(* IEC 61131-3 sources: Test002/ConveyorBelt/Class/VaranManager (part 2) *)

      7 : // all Varan_Base are ready with init
          if (s_ModuleList.ud_NrOfModules = 0) & (bEnableManagerWithNoModules = FALSE) then
            // penultimate call: if there are no clients => tell the hwcontrol to disable this
            To_HwControl.DisableVaranManager( ud_manager_number := VaranManagerNr
                                            , p_function_list   := #s_VMFunctions
                                            );
            State 		:= _NotInitialized;
          	ManagerOn := 0;                   //Disables Rt Task
          	bDisableCyTaskNoModules := TRUE;  //Disables Cy Task
          end_if;

    end_case;

    //trigger watchdog in init
    TriggerWatchdog();

  end_if;

  //increment our initcounter
  s_VaranManagerSettings.us_InitCounter += 1;

END_FUNCTION //VIRTUAL GLOBAL VaranManager::Init

//[#ENGLISH]
//=================================================================================================
//This function is called in PostScan by VaranManagerPostScan
//=================================================================================================
//[servers]	ManagerOn				:R		:state of Manager (On/Off)
//			RetryCounter			:W		:server counts retries
//			AsyVaranTime			:W		:time of asynchronous varan task
//[members]	s_CyHandles				:R		:structure to save Handles and thisp for cyclic update methodes
//			s_VaranTimes			:W		:structure for varan time measurement
//			us_UpdateOkCy			:R/W	:if variable = 1 then varan classes are called
//			p_ManagerStructure		:R		:pointer for manager structure (from OS)
//			s_VaranManagerSettings	:R/W	:structure for different varan settings
FUNCTION VIRTUAL GLOBAL VaranManager::CyWork
  VAR_INPUT
    EAX		              : UDINT;
  END_VAR
  VAR_OUTPUT
    state	    	        : UDINT;
  END_VAR
  VAR
    us_retry_counter	  : USINT;
    pHelp               : ^t_s_OneHandle;
    asyState            : UDINT;
    asyTimestamp        : UDINT;
  #ifndef VARAN_TIME_MEASUREMENT_DEACTIVATE
    ud_time				      : UDINT;
  #endif
    i				          	: UDINT;
    AsyReady            : BOOL;
    pHelpPostInit       : ^t_s_PostInitList;
  #ifdef VARAN_TIME_MEASUREMENT_SINGLE_OBJECTS
    ud_SingleTimeMark1  : UDINT;
    ud_SingleTimeMark2  : UDINT;
  #endif
  END_VAR

  //look if structur is ok, also check if cywork should be disabled due to no connected modules
  if ( p_ManagerStructure = NIL & b_PayloadSupport = false) | ( bDisableCyTaskNoModules = TRUE ) then
    return;
  end_if;

  //look if cyclic task is ready (executed)
  if b_PayloadSupport &
     pMultiVaran^.udVersion >= VM_MULTIVARAN_DOL_TIMING_AVAILABLE then

    MULTI_VARAN_iGetNodeProperty( hNodeHandle       := vmNodeHandle
                                , udPropertyId      := VM_PROP_TASK_STATE_ASY
                                , pudPropertyValue  := #asyState
                                );

    if asyState = TK_STATE_EXECUTING then
      AsyReady := FALSE;
    else
      AsyReady := TRUE;
    end_if;
  else
    AsyReady := (p_ManagerStructure^.sASY.ucHandshake and 16#10 ) <> 0;
  end_if;

#ifdef _LSL_TARGETARCH_ARM  // IO Image only needed for ARM  CPUs
#ifdef VARAN_iGetInputImage
  //look if manager is on or we are in post init phase (ManagerOn will be set in first realtime but we want to do something here in postinit)
  if ( ManagerOn = 1 ) | bPostInitActive = TRUE then
    if AsyReady then
      if b_IOImage then
        VARAN_iGetInputImage(VaranManagerNr, VARAN_DOL_ASY);
      end_if;
    end_if;
  end_if;
#endif
#endif

  // if there is a safety manager, we have to call it (but not from post init)
  if SafetyManagerThis & (bPostInitActive = FALSE) then
    SafetyManagerThis^.CyWork(0);
  end_if;

  //------------------------------------------------------------------------------------------------
  //first check Error
  if ( s_VaranManagerSettings.b_LogError = TRUE ) then
    LogError();
  end_if;

  // then check for rt log
  if bd_RtLog then
    if bd_RtLog.WatchdogTriggerFailed & (bd_RtLogged.WatchdogTriggerFailed = FALSE) then
#ifdef HWC_LogError
    HWC_LogError(this, "@0022 (VaranManager::CyWork) [SL] Error triggering the VaranManager Watchdog!");
#endif

      bd_RtLogged.WatchdogTriggerFailed := TRUE;
    end_if;

    if bd_RtLog.TimeSliceError & (bd_RtLogged.TimeSliceError = FALSE) then
#ifdef HWC_LogError
      HWC_LogError(this,"@019A (VaranManager::CyWork) Timeslice Error! Manager is set off!");
#endif

      bd_RtLogged.TimeSliceError := TRUE;
    end_if;

    bd_RtLog := 0;
  end_if;

#ifndef VARAN_TIME_MEASUREMENT_DEACTIVATE
  //measure time for cyclic
  ud_time := GetNsTime();
  s_VaranTimes.s_Cyclic.ud_CallTime := ( ud_time - s_VaranTimes.s_Cyclic.ud_Timemark ) / 1000;
  s_VaranTimes.s_Cyclic.ud_Timemark := ud_time;
#endif

  //check if we must disable a device
  if ( b_Disabledevice = TRUE ) then
    DisableDevice();
  end_if;

  //Update retry Counter
  if b_PayloadSupport &
     pMultiVaran^.udVersion >= VM_MULTIVARAN_VERSION_FULL_PAYLOAD_AVAILABLE  then
    MULTI_VARAN_iGetNodeProperty( hNodeHandle       := vmNodeHandle
                                , udPropertyId      := VM_PROP_GLOBAL_FAILED_ACCESS_COUNTER
                                , pudPropertyValue  := (#us_retry_counter)$^UDINT
                                );
  else
    us_retry_counter := p_ManagerStructure^.ucGlobalretryCounter;
  end_if;

  //look for change
  if ( us_retry_counter <> s_VaranManagerSettings.us_OldRetryCounter ) then

    //save on global counter
    RetryCounter += TO_USINT( us_retry_counter - s_VaranManagerSettings.us_OldRetryCounter );

    //save new counter
    s_VaranManagerSettings.us_OldRetryCounter := us_retry_counter;

    //update module retry counters cyclic
    if ( s_CyHandles.ud_NrOfHandles > 0 ) then

      //call all connected classes
      pHelp := #s_CyHandles.p_HandleList^[0];
      for i := 0 to s_CyHandles.ud_NrOfHandles - 1 do

        //call class
        pHelp^.p_This^.UpdateRetryCounter();

        //get pointer on next handle
        pHelp += sizeof(t_s_OneHandle);
      end_for;
    end_if;

    //update module retry counters cyclic
    if ( s_RtHandles.ud_NrOfHandles > 0 ) then

      //call all connected classes
      pHelp := #s_RtHandles.p_HandleList^[0];
      for i := 0 to s_RtHandles.ud_NrOfHandles - 1 do

        //call class
        pHelp^.p_This^.UpdateRetryCounter();

        //get pointer on next handle
        pHelp += sizeof(t_s_OneHandle);
      end_for;
    end_if;
  end_if;

  //look if manager is on or we are in post init phase (ManagerOn will be set in first realtime but we want to do something here in postinit)
  if ( ManagerOn = 1 ) | bPostInitActive = TRUE then

    //------------------------------------------------------------------------------------------------
    //look if cyclic task is ready (executed)
    if AsyReady = FALSE then
      s_VaranManagerSettings.us_NoCyclicUpdateCnt += 1;
      return;
    end_if;

#ifndef VARAN_TIME_MEASUREMENT_DEACTIVATE
    //------------------------------------------------------------------------------------------------
    //calculate cyclictime of varan task
    if b_PayloadSupport &
       pMultiVaran^.udVersion >= VM_MULTIVARAN_VERSION_FULL_PAYLOAD_AVAILABLE  then
      MULTI_VARAN_iGetNodeProperty( hNodeHandle       := vmNodeHandle
                                  , udPropertyId      := VM_PROP_ASY_TIME_UP_COUNTER
                                  , pudPropertyValue  := #asyTimestamp
                                  );
    else
      asyTimestamp := p_ManagerStructure^.sASY.uiTTUpCounter;
    end_if;

    if ( s_VaranTimes.s_AsyVaranTime.us_NotFirstRun	= 0 ) then

      //get counter of asy task
      s_VaranTimes.s_AsyVaranTime.ud_Timestamp := asyTimestamp;

      //start asy task
      if ( s_CyHandles.b_ExecuteDOL = TRUE ) then
        ExecuteDOL( VARAN_DOL_ASY );
      end_if;

      s_VaranTimes.s_AsyVaranTime.us_NotFirstRun := 1;
      return;
    end_if;

    //calculate ASY Time
    s_VaranTimes.s_AsyVaranTime.ud_ActUsageRate := asyTimestamp - s_VaranTimes.s_AsyVaranTime.ud_Timestamp;
    s_VaranTimes.s_AsyVaranTime.ud_Timestamp    := asyTimestamp;

    //look for maximum value
    if ( s_VaranTimes.s_AsyVaranTime.ud_ActUsageRate > s_VaranTimes.s_AsyVaranTime.ud_MaxUsageRate ) then
      s_VaranTimes.s_AsyVaranTime.ud_MaxUsageRate := s_VaranTimes.s_AsyVaranTime.ud_ActUsageRate;
    end_if;

    //save on server
    AsyVaranTime$UDINT := s_VaranTimes.s_AsyVaranTime.ud_ActUsageRate;
#endif

    //----------------------------------------------------------------------------------------------
    //hardware class handling

    // in post init we call only the modules which are logged in for post init
    if bPostInitActive then
      if PostInitModuleCnt then
        pHelpPostInit := #aPostInitList[0];
        for i := 0 to PostInitModuleCnt - 1 do

          //call class, if it's still not ready
          if pHelpPostInit^.p_This & pHelpPostInit^.b_CallMe then
            pHelpPostInit^.p_This^.UpdateCy();
          end_if;

          // set pointer on next this pointer
          pHelpPostInit += sizeof(t_s_PostInitList);
        end_for;
      end_if;
    else
      //look if we have classes
      if ( s_CyHandles.ud_NrOfHandles > 0 ) then

        //call all connected classes
        pHelp := #s_CyHandles.p_HandleList^[0];
        for i := 0 to s_CyHandles.ud_NrOfHandles - 1 do

#ifdef VARAN_TIME_MEASUREMENT_SINGLE_OBJECTS
          ud_SingleTimeMark1 := OS_READMICROSEC();
#endif

          //call class
          pHelp^.p_This^.UpdateCy();

#ifdef VARAN_TIME_MEASUREMENT_SINGLE_OBJECTS
          ud_SingleTimeMark2 := OS_READMICROSEC();
          pHelp^.TimeMeasuring.ud_ActTime := ud_SingleTimeMark2 - ud_SingleTimeMark1;

          if pHelp^.TimeMeasuring.ud_ActTime > pHelp^.TimeMeasuring.ud_MaxTime then
            pHelp^.TimeMeasuring.ud_MaxTime := pHelp^.TimeMeasuring.ud_ActTime;
          end_if;

          if pHelp^.TimeMeasuring.ud_ActTime < pHelp^.TimeMeasuring.ud_MinTime then
            pHelp^.TimeMeasuring.ud_MinTime := pHelp^.TimeMeasuring.ud_ActTime;
          end_if;
#endif

          //get pointer on next handle
          pHelp += sizeof(t_s_OneHandle);
        end_for;
      end_if;
    end_if;

    //start asy task
    if ( s_CyHandles.b_ExecuteDOL = TRUE ) then
      ExecuteDOL( VARAN_DOL_ASY );
    end_if;

  //------------------------------------------------------------ Client Instructions --------------------------------------------------------|
  //                                                                                                                                         V
    //DPRAM data handling
    if ( IsAlsoClient & p_ManagerClientSpace <> NIL ) then

      // copy data to ram
      // ->WRITE<-
      To_Stdlib.MemCpy( dest := #p_ASYDataWrite^.a_Data[0],     // Mem for p_ASYDataWrite is reserved in VaranManager2
                        source := AsyWriteData.pSDOData,        // Mem for AsyWriteData is reserved in VaranManager2
                        size := SafetyAsyMemWrite$UDINT
                      );

      // copy user data from application memory
      if UserObjectData.pAsyWriteData then
        To_Stdlib.MemCpy( dest := #p_ASYDataWrite^.a_Data[0] + SafetyAsyMemWrite,
                          source := UserObjectData.pAsyWriteData,
                          size := UserObjectData.udAsyWriteLength
                        );
    end_if;

      if (SafetyAsyMemWrite$UDINT + UserObjectData.udAsyWriteLength) > sizeof(UDINT) then
          To_Stdlib.MemCpy( dest    := p_ManagerClientSpace + VM_CLIENT_ASY_WR_OFFSET + sizeof(UDINT)
                          , source  := p_ASYDataWrite + sizeof(UDINT)
                          , size    := SafetyAsyMemWrite$UDINT + UserObjectData.udAsyWriteLength - sizeof(UDINT)
                          );
      end_if;

      //copy the first 4 bytes to DPRAM (to switch the shift buffer at the right moment)
      ((p_ManagerClientSpace + VM_CLIENT_ASY_WR_OFFSET)$^UDINT)^  := (p_ASYDataWrite$^UDINT)^;

      // copy read data to allocated space
      // ->READ<-
      if (SafetyAsyMemRead$UDINT + UserObjectData.udAsyReadLength) > sizeof(UDINT) then
        To_Stdlib.MemCpy( dest    := #p_ASYDataRead^.a_Data[0] + sizeof(UDINT)
                        , source  := p_ManagerClientSpace + VM_CLIENT_ASY_RD_OFFSET + sizeof(UDINT)
                        , size    := SafetyAsyMemRead$UDINT + UserObjectData.udAsyReadLength - sizeof(UDINT)
                        );
            end_if;

      //copy the first 4 bytes out of DPRAM (to switch the shift buffer at the right moment)
      (p_ASYDataRead$^UDINT)^ := ((p_ManagerClientSpace + VM_CLIENT_ASY_RD_OFFSET)$^UDINT)^;

      // copy data to application memory
      To_Stdlib.MemCpy( dest    := AsyReadData.pSDOData,
                        source  := #p_ASYDataRead^.a_Data[0],
                        size    := SafetyAsyMemRead$UDINT
                      );

      // copy user data to application memory
      if UserObjectData.pAsyReadData then
        To_Stdlib.MemCpy( dest    := UserObjectData.pAsyReadData,
                          source  := #p_ASYDataRead^.a_Data[0] + SafetyAsyMemRead,
                          size    := UserObjectData.udAsyReadLength
                        );
      end_if;

    end_if;
//------------------------------------------------------------ Client Instructions --------------------------------------------------------^
//                                                                                                                                         |
  end_if;

#ifndef VARAN_TIME_MEASUREMENT_DEACTIVATE
  //get cyclic time
  ud_time := GetNsTime();
  s_VaranTimes.s_Cyclic.ud_ActTime := ( ud_time - s_VaranTimes.s_Cyclic.ud_Timemark ) /1000;

  //get maximal time
  if ( s_VaranTimes.s_Cyclic.ud_ActTime > s_VaranTimes.s_Cyclic.ud_MaxTime ) then
    s_VaranTimes.s_Cyclic.ud_MaxTime := s_VaranTimes.s_Cyclic.ud_ActTime;
      end_if;
#endif

  State := READY;

END_FUNCTION //VIRTUAL GLOBAL VaranManager::CyWork
//[#ENGLISH]
//=================================================================================================
//Normal Rt - Funktion for VaranManager_Base
//=================================================================================================
//[servers]	ManagerOn				:R		:marks VaranManager as valid / ok
//			IsoVaranTime			:W		:time of isochronous varan task
//[members]	s_RtHandles				:R		:structure to save Handles and thisp for realtime update methodes
//			s_VaranTimes			:W		:structure for varan time measurement
//			us_UpdateOkRt			:R/W	:if variable = 1 then varan classes are called
//			p_ManagerStructure		:R		:pointer for manager structure (from OS)
//			s_VaranManagerSettings	:R/W	:structure for different varan settings
//			p_SyncOut				:R		:pointer to Varan sync out
//			p_SyncData				:R		:pointer to sync data object
FUNCTION VIRTUAL GLOBAL VaranManager::RtWork
  VAR_INPUT
    EAX		                    : UDINT;
  END_VAR
  VAR_OUTPUT
    state	    	              : UDINT;
  END_VAR
  VAR
    i			                    : UDINT;
    pHelp                     : ^t_s_OneHandle;
  #ifndef VARAN_TIME_MEASUREMENT_DEACTIVATE
    ud_time				            : UDINT;
    ud_IsoDuration            : UDINT;
  #endif
    ud_IsoState               : UDINT;
    systemProperty            : LSL_PROPERTY_VALUE_PAIR;
    us_newFrameCountThreshold : USINT;
    us_ControlStatus          : USINT;

  #ifdef VARAN_TIME_MEASUREMENT_SINGLE_OBJECTS
    ud_SingleTimeMark1        : UDINT;
    ud_SingleTimeMark2        : UDINT;
  #endif
  END_VAR

  //------------------------------------------------------------------------------------------------
  //if manager is not initialized
  if ( ManagerOn = -1 ) then

    // activate sync out for iso buffer
    if IsAlsoClient then  // ----------------------------------------------------------------------------------------------------

      // wait until hw-classes are synchrony
      if s_VMFunctions.b_HWClassSynchron = FALSE then

        //first trigger watchdog
        if ( b_RtDebug | ops.tAbsolute - s_VaranManagerSettings.ud_WatchdogTimemark > VM_WATCHDOG_TRIGGER_TIME ) then

          s_VaranManagerSettings.ud_WatchdogTimemark := ops.tAbsolute;
          TriggerWatchdog();			//trigger watchdog on varan Manager (local)
        end_if;
        return;
      end_if;

      // after this step, it's not necessary to check framecounter in hw_control anymore
      s_VMFunctions.b_OverrideFrameCheck := TRUE;

      // if superior system is slower, start with the sync after next
      if SuperiorSystemTime > VaranManagerTime then

        if b_PayloadSupport &
          pMultiVaran^.udVersion >= VM_MULTIVARAN_VERSION_FULL_PAYLOAD_AVAILABLE  then
          MULTI_VARAN_iGetNodeProperty( hNodeHandle       := vmNodeHandle
                                      , udPropertyId      := VM_PROP_PLL_SYNC_TIME_FRAME_COUNTER
                                      , pudPropertyValue  := (#us_newFrameCountThreshold)$^UDINT
                                      );
          us_newFrameCountThreshold += 2;
        else
          us_newFrameCountThreshold := p_ManagerPll^.ucSyncTimeFrameCounter + 2;
        end_if;

        p_SyncOut^.ucFrameCountThreshold := us_newFrameCountThreshold;
        p_SyncOutISOSwitch^.ucFrameCountThreshold := us_newFrameCountThreshold;

      else
      // otherwise don't use syncframecounter
        ucIsoSwitchTemp     := ucIsoSwitchTemp    AND 2#11111101;
        ucVaranManagerTemp  := ucVaranManagerTemp AND 2#11111101;
      end_if;

      p_SyncOutISOSwitch^.ucControlStatus := ucIsoSwitchTemp;

      // Write p_SyncOutISOSwitch
      if b_PayloadSupport &
          pMultiVaran^.udVersion >= VM_MULTIVARAN_VERSION_GET_SYSTEM_PROPERTY_AVAILABLE then
        MULTI_VARAN_ICONFIGUREPLLSYNCOUT( hManagerNodeHandle    := vmNodeHandle
                                        , udSyncOutId           := VM_CLIENT_ISO_SWITCH_ID
                                        , udPeriodMultiplier    := p_SyncOutISOSwitch^.ucPeriodMultiplier
                                        , udFrameCountThreshold := p_SyncOutISOSwitch^.ucFrameCountThreshold
                                        , udControlStatus       := p_SyncOutISOSwitch^.ucControlStatus
                                        );
      end_if;

      // activate sync out for varan manager (bit0 = 1)
      p_SyncOut^.ucControlStatus := ucVaranManagerTemp;
    else
      // activate sync out for varan manager (bit0 = 1)
      p_SyncOut^.ucControlStatus := 1;

    end_if; // if IsAlsoClient // ----------------------------------------------------------------------------------------------------

      // Always write sync out, cannot directly be written with payload support
    if b_PayloadSupport &
       pMultiVaran^.udVersion >= VM_MULTIVARAN_VERSION_GET_SYSTEM_PROPERTY_AVAILABLE  then
      MULTI_VARAN_ICONFIGUREPLLSYNCOUT( hManagerNodeHandle    := vmNodeHandle
                                      , udSyncOutId           := VM_SYNC_OUT_ID
                                      , udPeriodMultiplier    := p_SyncOut^.ucPeriodMultiplier
                                      , udFrameCountThreshold := p_SyncOut^.ucFrameCountThreshold
                                      , udControlStatus       := p_SyncOut^.ucControlStatus
                                      );
    end_if;

    //set manager on
    ManagerOn                             := 1;

    //to wait until we must be sync
    s_VaranManagerSettings.us_Wait4Sync   := 3;

    //to wait for Rtwork, we must be sync
    s_VaranManagerSettings.us_Wait4RtWork := 7;

    us_RtStep := _Wait4Sync;
    return;
  end_if;

  //------------------------------------------------------------------------------------------------
  //check if manager on
  if ( ManagerOn <> 1 ) then
    return;
  end_if;

  //first trigger watchdog
  if ( b_RtDebug | ops.tAbsolute - s_VaranManagerSettings.ud_WatchdogTimemark > VM_WATCHDOG_TRIGGER_TIME ) then

    s_VaranManagerSettings.ud_WatchdogTimemark := ops.tAbsolute;
    TriggerWatchdog();			//trigger watchdog on varan Manager (local)

    // trigger watchdog on clients (only if vmc is waiting for beeing synchron)
    if TriggerClientWD then

      if b_PayloadSupport &
         pMultiVaran^.udVersion >= VM_MULTIVARAN_VERSION_FULL_PAYLOAD_AVAILABLE  then
        MULTI_VARAN_iTriggerWatchdog( hManagerNodeHandle  := vmNodeHandle
                                    , udWatchdogType      := LSL_WD_TYPE_CLIENT
                                    );
      else

#ifdef VARAN_iTriggerClientWd
        VARAN_iTriggerClientWd(VaranManagerNr);
#endif
      end_if;
    end_if;
  end_if;

#ifdef _LSL_TARGETARCH_ARM  // IO Image only needed for ARM  CPUs
#ifdef VARAN_iGetInputImage
  if b_IOImage then
    VARAN_iGetInputImage(VaranManagerNr, VARAN_DOL_ISO);
  end_if;
#endif
#endif

  // Payload Support
  if b_PayloadSupport &
     pMultiVaran^.udVersion >= VM_MULTIVARAN_VERSION_FULL_PAYLOAD_AVAILABLE then
      //set frame counter in Sync data object and trigger client watchdogs
      MULTI_VARAN_iIncrementSyncCounter(hManagerNodeHandle := vmNodeHandle);
  else
    //set frame counter in Sync data object and trigger client watchdogs
    p_SyncData^.us_FrameCounter := p_SyncData^.us_FrameCounter + 1;
  end_if;

  //------------------------------------------------------------------------------------------------
  //look which step we have
  case ( us_RtStep ) of
//**********************************************************************************************************************************************************
    _Wait4Sync:		//wait some ticks (to be synchron)
      //look for either sync counter is zero or pll is locked and device delay time is compensated (if we use VMC)
      if ( s_VaranManagerSettings.us_Wait4Sync = 0 ) then
        us_RtStep := _InitVaranManager;
        return;
      elsif IsAlsoClient then

        // Read Pll Status Register
        if b_PayloadSupport &
           pMultiVaran^.udVersion >= VM_MULTIVARAN_VERSION_FULL_PAYLOAD_AVAILABLE  then
          MULTI_VARAN_iGetNodeProperty( hNodeHandle       := vmNodeHandle
                                      , udPropertyId      := VM_PROP_PLL_STATUS_REGISTER
                                      , pudPropertyValue  := (#us_ControlStatus)$^UDINT
                                      );
        else

          us_ControlStatus := p_ManagerPll^.ucControlStatus;
        end_if;

        if (((us_ControlStatus AND 2#0101) <> 2#0101) | (s_VMFunctions.b_HWClassSynchron = FALSE)) then
          // do countdown just after we got pll synchrony
          return;
        end_if;
      end_if;

      s_VaranManagerSettings.us_Wait4Sync -= 1;

//**********************************************************************************************************************************************************
    _InitVaranManager:		//Init Varan Manager (OS)

      if b_PayloadSupport &
         pMultiVaran^.udVersion >= VM_MULTIVARAN_VERSION_FULL_PAYLOAD_AVAILABLE  then // ---------------------------------------------------------------------------------

        //call init of OS to init varan command list and start varan bus
        // (Replaces VARAN_iInitApp)

        //Only set system properties once per system
        if (bSetSystemProperties = TRUE) then

          systemProperty.udPropertyId     := SYS_PROP_OPERATIONAL_STATE;
          systemProperty.udPropertyValue  := OP_STATE_POST_INIT;
          MULTI_VARAN_iSetSystemProperties( udPropertyCount       := 1
                                          , psPropertyValuePairs  := #systemProperty
                                          );
        end_if;

#ifndef VARAN_TIME_MEASUREMENT_DEACTIVATE
        //get iso counter of FPGA to calculate ISO Time
        MULTI_VARAN_iGetIsoDuration ( hManagerNodeHandle  := vmNodeHandle
                                    , pudIsoDurationNs    := #s_VaranTimes.s_IsoVaranTime.ud_Timestamp
                                    );
#endif

        //get old retry counter
        MULTI_VARAN_iGetNodeProperty( hNodeHandle       := vmNodeHandle
                                    , udPropertyId      := VM_PROP_GLOBAL_FAILED_ACCESS_COUNTER
                                    , pudPropertyValue  := (#s_VaranManagerSettings.us_OldRetryCounter)$^UDINT
                                    );
      else  // if b_PayloadSupport then // ---------------------------------------------------------------------------------

        //call init of OS to init varan command list and start varan bus
        if pVaran then
          VARAN_iInitApp( VaranManagerNr );
        end_if;

#ifndef VARAN_TIME_MEASUREMENT_DEACTIVATE
      //get iso counter of FPGA to calculate ISO Time
      s_VaranTimes.s_IsoVaranTime.ud_Timestamp := p_ManagerStructure^.sISO.uiReserved2;
#endif

        //get old retry counter
        s_VaranManagerSettings.us_OldRetryCounter := p_ManagerStructure^.ucGlobalretryCounter;
      end_if; // if b_PayloadSupport then // ---------------------------------------------------------------------------------

      //start iso task first time
      ExecuteDOL( VARAN_DOL_ISO );

      //next step
      us_RtStep := _Wait4RtWork;

//**********************************************************************************************************************************************************
    _Wait4RtWork://wait for RtWork -> syncs, which are enabled in _InitVaranManager are send now

      if b_PayloadSupport &
         pMultiVaran^.udVersion >= VM_MULTIVARAN_DOL_TIMING_AVAILABLE then
      //look if realtime of VaranManager has finished
        MULTI_VARAN_iCheckIsoState( hManagerNodeHandle := vmNodeHandle
                                  , pudIsoState        := #ud_IsoState
                                  );

        if ud_IsoState = TK_STATE_EXECUTING then
          TRACE_RtOverlap();
          return;
        end_if;
      else
          //look if realtime of VaranManager has finished
        if ( ( p_ManagerStructure^.sISO.ucHandshake and 16#10 ) = 0 ) then
          TRACE_RtOverlap();
          return;
        end_if;
      end_if;

      if s_VaranManagerSettings.us_Wait4RtWork = 0 then
#ifndef VARAN_TIME_MEASUREMENT_DEACTIVATE
        //take timestamp
        if b_PayloadSupport &
           pMultiVaran^.udVersion >= VM_MULTIVARAN_VERSION_FULL_PAYLOAD_AVAILABLE  then
          MULTI_VARAN_iGetTimeUpCounter( hManagerNodeHandle := vmNodeHandle
                                       , pudTimeUpCounterNs  := #s_VaranTimes.s_Realtime.ud_Timemark
                                       );
        else
        s_VaranTimes.s_Realtime.ud_Timemark := p_ManagerStructure^.uiTUpCounter;
        end_if;

        Max_RtCallTime := 0;
        Min_RtCallTime := 16#FFFF_FFFF;
        Max_RtTime := 0;
        Min_RtTime := 16#FFFF_FFFF;
#endif
        us_RtStep := _RtWork;
      else
        ExecuteDOL( VARAN_DOL_ISO );  // Don't Execute when switching to _RtWork, UpDateRtPostscan takes over this call
      end_if;

      s_VaranManagerSettings.us_Wait4RtWork -= 1;

//**********************************************************************************************************************************************************
    _RtWork://normal RtWork

#ifndef VARAN_TIME_MEASUREMENT_DEACTIVATE
      //get time in ns
      if b_PayloadSupport &
         pMultiVaran^.udVersion >= VM_MULTIVARAN_VERSION_FULL_PAYLOAD_AVAILABLE  then
        MULTI_VARAN_iGetTimeUpCounter( hManagerNodeHandle := vmNodeHandle
                                     , pudTimeUpCounterNs := #ud_time
                                     );
      else
        ud_time := p_ManagerStructure^.uiTUpCounter;
      end_if;

      //get call time
      Act_RtCallTime := ( ud_time - s_VaranTimes.s_Realtime.ud_Timemark ) / 1000;
      s_VaranTimes.s_Realtime.ud_Timemark := ud_time;

      //look for maximum
      if ( Act_RtCallTime > Max_RtCallTime ) then
        Max_RtCallTime := Act_RtCallTime;
      end_if;

      //look for minimum
      if ( Act_RtCallTime < Min_RtCallTime ) then
        Min_RtCallTime := Act_RtCallTime;
      end_if;

      //calculate ISO Time
      if b_PayloadSupport &
         pMultiVaran^.udVersion >= VM_MULTIVARAN_DOL_TIMING_AVAILABLE then
        MULTI_VARAN_iGetIsoDuration ( hManagerNodeHandle  := vmNodeHandle
                                    , pudIsoDurationNs    := #s_VaranTimes.s_IsoVaranTime.ud_ActUsageRate
                                    );
      else
        ud_IsoDuration := p_ManagerStructure^.sISO.uiReserved2;

        s_VaranTimes.s_IsoVaranTime.ud_ActUsageRate := ud_IsoDuration - s_VaranTimes.s_IsoVaranTime.ud_Timestamp;
        s_VaranTimes.s_IsoVaranTime.ud_Timestamp := ud_IsoDuration;
      end_if;

      //look for maximum value
      if ( s_VaranTimes.s_IsoVaranTime.ud_ActUsageRate > IsoVaranTimeMax ) then
        if s_VaranTimes.s_IsoVaranTime.us_NotFirstRun = 0 then
          s_VaranTimes.s_IsoVaranTime.us_NotFirstRun := 1;
        else
          IsoVaranTimeMax := s_VaranTimes.s_IsoVaranTime.ud_ActUsageRate;
        end_if;
      end_if;

      //save on server
      IsoVaranTime$UDINT := s_VaranTimes.s_IsoVaranTime.ud_ActUsageRate;
#endif

      if b_PayloadSupport &
         pMultiVaran^.udVersion >= VM_MULTIVARAN_DOL_TIMING_AVAILABLE then
      //look if realtime of VaranManager has finished
        MULTI_VARAN_iCheckIsoState( hManagerNodeHandle := vmNodeHandle
                                  , pudIsoState        := #ud_IsoState
                                  );

        if ud_IsoState = TK_STATE_EXECUTING then
          TRACE_RtOverlap();
          return;
        end_if;
      else
          //look if realtime of VaranManager has finished
        if ( ( p_ManagerStructure^.sISO.ucHandshake and 16#10 ) = 0 ) then
          TRACE_RtOverlap();
          return;
        end_if;
      end_if;

      //----------------------------------------------------------------------------------------------
      //hardware class handling

      //look if we have classes
      if ( s_RtHandles.ud_NrOfHandles > 0 ) then

        //call all connected classes
        pHelp := #s_RtHandles.p_HandleList^[0];

        // faster from 1 to number than from 0 to number-1
        for i := 1 to s_RtHandles.ud_NrOfHandles do
#ifdef VARAN_TIME_MEASUREMENT_SINGLE_OBJECTS
          ud_SingleTimeMark1 := OS_READMICROSEC();
#endif

          //call class
          pHelp^.p_This^.UpdateRt();

#ifdef VARAN_TIME_MEASUREMENT_SINGLE_OBJECTS
          ud_SingleTimeMark2 := OS_READMICROSEC();
          pHelp^.TimeMeasuring.ud_ActTime := ud_SingleTimeMark2 - ud_SingleTimeMark1;

          if pHelp^.TimeMeasuring.ud_ActTime > pHelp^.TimeMeasuring.ud_MaxTime then
            pHelp^.TimeMeasuring.ud_MaxTime := pHelp^.TimeMeasuring.ud_ActTime;
          end_if;

          if pHelp^.TimeMeasuring.ud_ActTime < pHelp^.TimeMeasuring.ud_MinTime then
            pHelp^.TimeMeasuring.ud_MinTime := pHelp^.TimeMeasuring.ud_ActTime;
          end_if;
#endif

          //get pointer on next handle
          pHelp += sizeof(t_s_OneHandle);
        end_for;
      end_if;

  //------------------------------------------------------------ Client Instructions --------------------------------------------------------|
  //                                                                                                                                         V
      //copy client data out of DPRAM, if we are synchrony
      if ( IsAlsoClient & p_ManagerClientSpace <> NIL ) then

        //--------------------------------------------------------------------------------------------------------------------------------------
        if bPdoCopyDisable = false then  // PDO data are copied automatic
          // copy data to application memory
          if pIsoReadSafetyData then
            To_Stdlib.MemCpy( dest    := pIsoReadSafetyData,
                              source 	:= p_ManagerClientSpace + VM_CLIENT_ISO_RD_OFFSET,
                              size    := SafetyIsoMemRead$UDINT + VM_CLIENT_HEADER_SIZE
                            );
          end_if;
        else
          // copy data to application memory
          if pIsoReadSafetyData then
            To_Stdlib.MemCpy( dest    := pIsoReadSafetyData,
                              source  := p_ManagerClientSpace + VM_CLIENT_ISO_RD_OFFSET,
                              size    := sizeof(t_VMC_Header) + sizeof(t_VMC_Safety_Header_TDO)
                              );
          end_if;
        end_if;

        // copy user PDO data from application to manager DPRAM
        if UserObjectData.pIsoReadData then
          To_Stdlib.MemCpy( dest    := UserObjectData.pIsoReadData,
                            source  := p_ManagerClientSpace + VM_CLIENT_ISO_RD_OFFSET + SafetyIsoMemRead + VM_CLIENT_HEADER_SIZE,
                            size    := UserObjectData.udIsoReadLength
                          );
        end_if;
      //--------------------------------------------------------------------------------------------------------------------------------------

      end_if;

  //------------------------------------------------------------ Client Instructions --------------------------------------------------------^
//**********************************************************************************************************************************************************
  end_case;

  State := READY;

END_FUNCTION //VIRTUAL GLOBAL VaranManager::RtWork

//[#ENGLISH]
//=================================================================================================
//Function to add a realtime or cyclic task to VaranManager
//=================================================================================================
//[server]	State					:R		:State of class
//[members]	s_RtHandles				:R/W	:structure to save Handles and thisp for realtime update methodes
//			s_CyHandles				:R/W	:structure to save Handles and thisp for cyclic update methodes
//[locals]	p_one_handle			:W/R	:pointer to next handle in list
//[>ud_dol_type] type of DOL list( Realtime = 3, cyclic = 4 )
//[>p_this] Thispointer of connected varan class
FUNCTION VIRTUAL GLOBAL VaranManager::AddVaranTask
  VAR_INPUT
    ud_dol_type 	: UDINT;
    p_this 	      : ^void;
    callOptions 	: USINT;
  END_VAR
  VAR
    p_one_handle	: ^t_s_OneHandle;
  END_VAR

  //look if we have a thispointer
  if (p_this <> NIL) then

    //------------------------------------------------------------------------------------------------
    //realtime
    if ( ud_dol_type = VARAN_DOL_ISO ) then
      IF callOptions AND CALL_OPTION_RT_PRESCAN THEN
        //is list full
        if ( s_RtHandles.ud_NrOfHandles = s_RtHandles.ud_MaxHandles ) then

          //extend list
          ExtendHandleList( ud_dol_type := VARAN_DOL_ISO );

          //if an error occured return
          if ( State <> _ClassOk ) then
            return;
          end_if;
        end_if;

        //set pointer to next free handle entry
        p_one_handle 			    := s_RtHandles.p_HandleList + ( s_RtHandles.ud_NrOfHandles * sizeof( t_s_OneHandle ) );
        p_one_handle^.p_This 	:= p_this$p_VaranBase;

#ifdef VARAN_TIME_MEASUREMENT_SINGLE_OBJECTS
        p_one_handle^.TimeMeasuring.ud_MinTime := 16#FFFFFFFF;
        _GetObjName( p_this$pVirtualBase, #p_one_handle^.TimeMeasuring.aObjname[0] );
#endif

        //increase number of handles
        s_RtHandles.ud_NrOfHandles += 1;
      END_IF;

      IF callOptions AND CALL_OPTION_RT_POSTSCAN THEN
        //is list full
        if ( s_RtPostScanHandles.ud_NrOfHandles = s_RtPostScanHandles.ud_MaxHandles ) then

          //extend list
          ExtendHandleList( ud_dol_type := VARAN_DOL_ISO, callOptions := CALL_OPTION_RT_POSTSCAN );

          //if an error occured return
          if ( State <> _ClassOk ) then
            return;
          end_if;
        end_if;

        //set pointer to next free handle entry
        p_one_handle 			    := s_RtPostScanHandles.p_HandleList + ( s_RtPostScanHandles.ud_NrOfHandles * sizeof( t_s_OneHandle ) );
        p_one_handle^.p_This 	:= p_this$p_VaranBase;

#ifdef VARAN_TIME_MEASUREMENT_SINGLE_OBJECTS
        p_one_handle^.TimeMeasuring.ud_MinTime := 16#FFFFFFFF;
        _GetObjName( p_this$pVirtualBase, #p_one_handle^.TimeMeasuring.aObjname[0] );
#endif

        //increase number of handles
        s_RtPostScanHandles.ud_NrOfHandles += 1;
      END_IF;
    //------------------------------------------------------------------------------------------------
    //cyclic
    elsif ( ud_dol_type = VARAN_DOL_ASY ) then

      //is list full
      if ( s_CyHandles.ud_NrOfHandles = s_CyHandles.ud_MaxHandles ) then

        //extend list
        ExtendHandleList( ud_dol_type := VARAN_DOL_ASY );

        //is an error occured
        if ( State <> _ClassOk ) then
          return;
        end_if;
      end_if;

      //set pointer to next free handle entry
      p_one_handle 			    := s_CyHandles.p_HandleList + ( s_CyHandles.ud_NrOfHandles * sizeof( t_s_OneHandle ) );
      p_one_handle^.p_This 	:= p_this$p_VaranBase;

#ifdef VARAN_TIME_MEASUREMENT_SINGLE_OBJECTS
        p_one_handle^.TimeMeasuring.ud_MinTime := 16#FFFFFFFF;
        _GetObjName( p_this$pVirtualBase, #p_one_handle^.TimeMeasuring.aObjname[0] );
#endif

      //increase number of handles
      s_CyHandles.ud_NrOfHandles += 1;
    end_if;
  end_if;

END_FUNCTION //VIRTUAL GLOBAL VaranManager::AddVaranTask

//[#ENGLISH]
//=================================================================================================
//Function to add a read data object to varan Manager and install a varan task
//=================================================================================================
//[members] s_CyHandles			:W		:structure to save Handles and thisp for cyclic update methodes
//[locals]	ud_command			:W/R	:to save right command for DO
//[>p_us_position_info]pointer to position info( first byte is length)
//[>ud_dol_type] type of DOL list( 1=direct access, 2=IRQ, 3=realtime, 4=cyclic )
//[>p_ud_handle]pointer to variable to set right handle
//[>ud_address] Address of data object
//[>ud_length] Length of data object
//[>p_ud_data] pointer to variable to get pointer to data
//[>ud_type]0=control area, 1=memory area
//[<sd_retval] 0=OK, negative=error (look lsl_st_varan.h)
FUNCTION VIRTUAL GLOBAL VaranManager::AddRdDO
VAR_INPUT
  p_us_position_info	: ^USINT;
  ud_dol_type		    	:  UDINT;
  p_ud_handle		    	: ^UDINT;
  ud_address		    	:  UDINT;
  ud_length			      :  UDINT;
  p_ud_data		      	: ^UDINT;
  ud_type			       	:  UDINT;
END_VAR
VAR_OUTPUT
  sd_retval			      :  DINT;
END_VAR
VAR
  ud_command		    	:  UDINT;
  TempMem             :  UDINT;
END_VAR

#ifdef VM_DEBUG_PAYLOAD
  // Payload not supported
  if b_PayloadSupport then
   // This method is not supporded with Payload support
    ((0)$^USINT)^ := 0;
  end_if;
#endif
  // if there is no VARAN Interface available, we would crash at the VARAN_iAddDOToDOL call
  if pVaran = NIL then
    sd_retval := VARANMANAGER_DRIVER_NOT_EXISTS;
    return;
  end_if;

  //look which type it is
  if ( ud_type AND 1) = 1 then
    ud_command := VARAN_CMD_MEMORY_READ;		//memory area
  else
    ud_command := VARAN_CMD_CONTROL_READ;		//control area
  end_if;

  //look if we must execute Cyclic DOL list
  if ( ud_dol_type = VARAN_DOL_ASY ) then
    s_CyHandles.b_ExecuteDOL := TRUE;			//set flag to execut Dol list
  end_if;

  //Install Varan data object
  sd_retval := VARAN_iAddDOToDOL	( uiManager			  := VaranManagerNr
                                  , pucNode			    := p_us_position_info
                                  , uiDOLType 		  := ud_dol_type
                                  , puiDOHandle		  := p_ud_handle
                                  , uiCmd				    := ud_command
                                  , uiAddressRead		:= ud_address
                                  , uiLengthRead		:= ud_length
                                  , pucRead			    := p_ud_data
                                  , uiAddressWrite	:= 0
                                  , uiLengthWrite		:= 0
                                  , pucWrite			  := NIL
                                  );

  //look if an error occured
  if ( sd_retval <> VARANMANAGER_OK ) then
    s_ErrorVaranManager.f_AddRdDO := SetVaranDOError( sd_Error 		  := sd_retval
                                                    , b_manager_off	:= TRUE
                                                    , b_log			    := TRUE
                                                    );
  else

    // check if the DO has a special priority
    if ud_type AND VM_PRIORITY_FILTER then
      AddToDOPriorityList(p_ud_handle^$^LSL_VARANFRAME, ud_type AND VM_PRIORITY_FILTER);
    end_if;

    // 32 Byte (Header) + 6 Byte (1 Byte Cmd, 4 Byte Addr, 1 Byte Len) + 1 Byte (Response) + n Byte (Load data read) + 0 to 3 Byte (compensate missalignment)
    TempMem := 32 + 6 + 1 + ud_length;
    if (TempMem MOD 4) then
      TempMem := TempMem + (4 - (TempMem MOD 4)); //increase memory, up to a value, which could be divided by 4
    end_if;

    case ud_dol_type of
    // **************************************************
      VARAN_DOL_DA:
        DPRAM_Used.DA_Rd    += TempMem;
        DOCounter.DA_Rd     += 1;
    // **************************************************
      VARAN_DOL_ISO:
        DPRAM_Used.ISO_Rd   += TempMem;
        DOCounter.ISO_Rd    += 1;
    // **************************************************
      VARAN_DOL_ASY:
        DPRAM_Used.ASY_Rd   += TempMem;
        DOCounter.ASY_Rd    += 1;
    // **************************************************
      VARAN_DOL_ADMIN:
        DPRAM_Used.Admin_Rd += TempMem;
        DOCounter.Admin_Rd  += 1;
    // **************************************************
      VARAN_DOL_IRQ:
        DPRAM_Used.IRQ_Rd   += TempMem;
        DOCounter.IRQ_Rd    += 1;
    end_case;

    DPRAM_Used.Total  += TempMem;
    DOCounter.Total   += 1;

  end_if;

END_FUNCTION //VIRTUAL GLOBAL VaranManager::AddRdDO

//[#ENGLISH]
//=================================================================================================
//Function to add a write data object to varan Manager and install a varan task
//=================================================================================================
//[members] s_CyHandles			:W		:structure to save Handles and thisp for cyclic update methodes
//[locals]	ud_command			:W/R	:to save right command for DO
//[>p_us_position_info]pointer to position info( first byte is length)
//[>ud_dol_type] type of DOL list( 1=direct access, 2=IRQ, 3=realtime, 4=cyclic )
//[>p_ud_handle]pointer to variable to set right handle
//[>ud_address] Address of data object
//[>ud_length] Length of data object
//[>p_ud_data] pointer to variable to get pointer to data
//[>ud_type]0=control area, 1=memory area
//[<sd_retval] 0=OK, negative=error (look lsl_st_varan.h)
FUNCTION VIRTUAL GLOBAL VaranManager::AddWrDO
VAR_INPUT
  p_us_position_info	  : ^USINT;
  ud_dol_type			      :  UDINT;
  p_ud_handle     			: ^UDINT;
  ud_address		      	:  UDINT;
  ud_length			        :  UDINT;
  p_ud_data			        : ^UDINT;
  ud_type			        	:  UDINT;
END_VAR
VAR_OUTPUT
  sd_retval			        :  DINT;
END_VAR
VAR
  ud_command		      	:  UDINT;
  TempMem               :  UDINT;
END_VAR

#ifdef VM_DEBUG_PAYLOAD
  // Payload not supported
  if b_PayloadSupport then
    // This method is not supporded with Payload support
    ((0)$^USINT)^ := 0;
  end_if;
#endif
  // if there is no VARAN Interface available, we would crash at the VARAN_iAddDOToDOL call
  if pVaran = NIL then
    sd_retval := VARANMANAGER_DRIVER_NOT_EXISTS;
    return;
  end_if;

  //look which type it is
  if ( ud_type AND 1) = 1 then
    ud_command := VARAN_CMD_MEMORY_WRITE;		//memory area
  else
    ud_command := VARAN_CMD_CONTROL_WRITE;		//control area
  end_if;

  //look if we must execute Cyclic DOL list
  if ( ud_dol_type = VARAN_DOL_ASY ) then
    s_CyHandles.b_ExecuteDOL := TRUE;			//set flag to execut Dol list
  end_if;

  //Install Varan data object
  sd_retval := VARAN_iAddDOToDOL	( uiManager			  := VaranManagerNr
                                  , pucNode			    := p_us_position_info
                                  , uiDOLType 		  := ud_dol_type
                                  , puiDOHandle		  := p_ud_handle
                                  , uiCmd				    := ud_command
                                  , uiAddressRead		:= 0
                                  , uiLengthRead		:= 0
                                  , pucRead			    := NIL
                                  , uiAddressWrite	:= ud_address
                                  , uiLengthWrite		:= ud_length
                                  , pucWrite			  := p_ud_data
                                  );

  //look if an error occured
  if ( sd_retval <> VARANMANAGER_OK ) then
    s_ErrorVaranManager.f_AddWrDO := SetVaranDOError	( sd_Error 		  := sd_retval
                                                      , b_manager_off	:= TRUE
                                                      , b_log			    := TRUE
                                                      );
  else

    // check if the DO has a special priority
    if ud_type AND VM_PRIORITY_FILTER then
      AddToDOPriorityList(p_ud_handle^$^LSL_VARANFRAME, ud_type AND VM_PRIORITY_FILTER);
    end_if;

    //32 Byte (Header) + 6 Byte (1 Byte Cmd, 4 Byte Addr, 1 Byte Len) + 1 Byte (Response) + n Byte (load data write) + 0 to 3 Byte (compensate missalignment)
    TempMem := 32 + 6 + 1 + ud_length;
    if (TempMem MOD 4) then
      TempMem := TempMem + (4 - (TempMem MOD 4)); //increase memory, up to a value, which could be divided by 4
    end_if;

    case ud_dol_type of
    // **************************************************
      VARAN_DOL_DA:
                    DPRAM_Used.DA_Wr    += TempMem;
                    DOCounter.DA_Wr     += 1;
    // **************************************************
      VARAN_DOL_ISO:
                    DPRAM_Used.ISO_Wr   += TempMem;
                    DOCounter.ISO_Wr    += 1;
    // **************************************************
      VARAN_DOL_ASY:
                    DPRAM_Used.ASY_Wr   += TempMem;
                    DOCounter.ASY_Wr    += 1;
    // **************************************************
      VARAN_DOL_ADMIN:
                    DPRAM_Used.Admin_Wr += TempMem;
                    DOCounter.Admin_Wr  += 1;
    // **************************************************
      VARAN_DOL_IRQ:
                    DPRAM_Used.IRQ_Wr   += TempMem;
                    DOCounter.IRQ_Wr    += 1;
      end_case;

      DPRAM_Used.Total  += TempMem;
      DOCounter.Total   += 1;
  end_if;

END_FUNCTION //VIRTUAL GLOBAL VaranManager::AddWrDO

//[#ENGLISH]
//=================================================================================================
//Function to add a read/write data object to varan manager and install a varan task
//=================================================================================================
//[members] s_CyHandles			:W		:structure to save Handles and thisp for cyclic update methodes
//[locals]	ud_command			:W/R	:to save right command for DO
//[>p_us_position_info]pointer to position info( first byte is length)
//[>ud_dol_type] type of DOL list( 1=direct access, 2=IRQ, 3=realtime, 4=cyclic )
//[>p_ud_handle] pointer to variable to set right handle
//[>ud_address_read] Address of read data object
//[>ud_length_read] Length of read data object
//[>p_ud_data_read] pointer to variable to get pointer to data
//[>ud_address_write] Address of write data object
//[>ud_length_write] Length of write data object
//[>p_ud_data_write] pointer to variable to get pointer to data
//[>ud_type]0=control area, 1=memory area
//[<sd_retval] 0=OK, negative=error (look lsl_st_varan.h)
FUNCTION VIRTUAL GLOBAL VaranManager::AddRdWrDO
  VAR_INPUT
    p_us_position_info	  : ^USINT;
    ud_dol_type			      :  UDINT;
    p_ud_handle			      : ^UDINT;
    ud_address_read		    :  UDINT;
    ud_length_read		    :  UDINT;
    p_ud_data_read		    : ^UDINT;
    ud_address_write	    :  UDINT;
    ud_length_write		    :  UDINT;
    p_ud_data_write		    : ^UDINT;
    ud_type				        :  UDINT;
  END_VAR
  VAR_OUTPUT
    sd_retval			        :  DINT;
  END_VAR
  VAR
    ud_command			      :  UDINT;
    TempMem               :  UDINT;
  END_VAR

#ifdef VM_DEBUG_PAYLOAD
  // Payload not supported
  if b_PayloadSupport then
    // This method is not supporded with Payload support
    ((0)$^USINT)^ := 0;
  end_if;
#endif
  // if there is no VARAN Interface available, we would crash at the VARAN_iAddDOToDOL call
  if pVaran = NIL then
    sd_retval := VARANMANAGER_DRIVER_NOT_EXISTS;
    return;
  end_if;

  //look which type it is
  if ( ud_type AND 1) = 1 then
    ud_command := VARAN_CMD_MEMORY_READ_WRITE;		//memory area
  else
    ud_command := VARAN_CMD_CONTROL_READ_WRITE;		//control area
  end_if;

  //look if we must execute Cyclic DOL list
  if ( ud_dol_type = VARAN_DOL_ASY ) then
    s_CyHandles.b_ExecuteDOL := TRUE;			//set flag to execut Dol list
  end_if;

  //Install Varan data object
  sd_retval := VARAN_iAddDOToDOL	( uiManager			  := VaranManagerNr
                                  , pucNode			    := p_us_position_info
                                  , uiDOLType 		  := ud_dol_type
                                  , puiDOHandle		  := p_ud_handle
                                  , uiCmd				    := ud_command
                                  , uiAddressRead		:= ud_address_read
                                  , uiLengthRead		:= ud_length_read
                                  , pucRead			    := p_ud_data_read
                                  , uiAddressWrite	:= ud_address_write
                                  , uiLengthWrite		:= ud_length_write
                                  , pucWrite			  := p_ud_data_write
                                  );

  //look if an error occured
  if ( sd_retval <> VARANMANAGER_OK ) then
    s_ErrorVaranManager.f_AddRdWrDO := SetVaranDOError	( sd_Error 		  := sd_retval
                                                        , b_manager_off	:= TRUE
                                                        , b_log			    := TRUE
                                                        );
  else

    // check if the DO has a special priority
    if ud_type AND VM_PRIORITY_FILTER then
      AddToDOPriorityList(p_ud_handle^$^LSL_VARANFRAME, ud_type AND VM_PRIORITY_FILTER);
    end_if;

    //32 Byte (Header) + 11 Byte (1 Byte Cmd, 4 Byte RdAddr, 1 Byte RdLen, 4 Byte WrAddr, 1 Byte WrLen) + 1 Byte (Response) + n Byte (load data read) + n Byte (load data write) + 0 to 3 Byte (compensate missalignment)
    TempMem := 32 + 11 + 1 + ud_length_read + ud_length_write;
    if (TempMem MOD 4) then
      TempMem := TempMem + (4 - (TempMem MOD 4)); //increase memory, up to a value, which could be divided by 4
    end_if;

    case ud_dol_type of
    // **************************************************
      VARAN_DOL_DA:
        DPRAM_Used.DA_RdWr    += TempMem;
        DOCounter.DA_RdWr     += 1;
    // **************************************************
      VARAN_DOL_ISO:
        DPRAM_Used.ISO_RdWr   += TempMem;
        DOCounter.ISO_RdWr    += 1;
    // **************************************************
      VARAN_DOL_ASY:
        DPRAM_Used.ASY_RdWr   += TempMem;
        DOCounter.ASY_RdWr    += 1;
    // **************************************************
      VARAN_DOL_ADMIN:
        DPRAM_Used.Admin_RdWr += TempMem;
        DOCounter.Admin_RdWr  += 1;
    // **************************************************
      VARAN_DOL_IRQ:
        DPRAM_Used.IRQ_RdWr   += TempMem;
        DOCounter.IRQ_RdWr    += 1;
    end_case;

    DPRAM_Used.Total  += TempMem;
    DOCounter.Total   += 1;
  end_if;

END_FUNCTION //VIRTUAL GLOBAL VaranManager::AddRdWrDO

//[#ENGLISH]
//=================================================================================================
//Function executes a data object list of VaranManager
//=================================================================================================
//[>ud_dol_type] type of DOL list( 1=direct access, 2=IRQ, 3=realtime, 4=cyclic )
//[<sd_retval] 0=OK, negative=error (look lsl_st_varan.h)
FUNCTION VIRTUAL GLOBAL VaranManager::ExecuteDOL
  VAR_INPUT
    ud_dol_type	      	: UDINT;
  END_VAR
  VAR_OUTPUT
    sd_retval	        	: DINT;
  END_VAR

  // Payload Support
  if b_PayloadSupport &
     pMultiVaran^.udVersion >= VM_MULTIVARAN_DOL_TIMING_AVAILABLE then

      //if we have a ARM CPU with payload, we have to set output image before we
#ifdef _LSL_TARGETARCH_ARM  // IO Image only needed for ARM  CPUs
#ifdef VARAN_iSetOutputImage
    if b_IOImage then
      VARAN_iSetOutputImage(VaranManagerNr, ud_dol_type);
    end_if;
#endif
#endif

    sd_retval := MULTI_VARAN_iExecuteDol( hManagerNodeHandle  := vmNodeHandle
                                        , udDolType           := ud_dol_type
                                        );

  else

    // if there is no VARAN Interface available, we would crash at the call
    if pVaran = NIL then
      sd_retval := VARANMANAGER_DRIVER_NOT_EXISTS;
      return;
    end_if;

    case ( ud_dol_type ) of

      VARAN_DOL_ISO:
#ifdef _LSL_TARGETARCH_ARM  // IO Image only needed for ARM  CPUs
#ifdef VARAN_iSetOutputImage
                      if b_IOImage then
                        VARAN_iSetOutputImage(VaranManagerNr, ud_dol_type);
                      end_if;
#endif
#endif

                      sd_retval := VARAN_iExecuteDOLISO( uiManager := VaranManagerNr );

      VARAN_DOL_ASY:
#ifdef _LSL_TARGETARCH_ARM  // IO Image only needed for ARM  CPUs
#ifdef VARAN_iSetOutputImage
                      if b_IOImage then
                        VARAN_iSetOutputImage(VaranManagerNr, ud_dol_type);
                      end_if;
#endif
#endif
                      sd_retval := VARAN_iExecuteDOLASY( uiManager := VaranManagerNr );

      VARAN_DOL_DA:	  sd_retval := VARAN_iExecuteDOLDA ( uiManager := VaranManagerNr );

      VARAN_DOL_IRQ:  sd_retval := VARAN_iExecuteDOLIRQ( uiManager := VaranManagerNr );
    end_case;
  end_if;

  //look if an error occurs
  if ( sd_retval <> VARANMANAGER_OK ) then
    s_ErrorVaranManager.f_ExecuteDOL := SetVaranDOError	( sd_Error 		  := sd_retval
                                                        , b_manager_off	:= TRUE
                                                        , b_log			    := TRUE
                                                        );
  end_if;

END_FUNCTION //VIRTUAL GLOBAL VaranManager::ExecuteDOL

//[#ENGLISH]
//=================================================================================================
//Function clears a data object list of VaranManager
//=================================================================================================
//[>ud_dol_type] Type of DOL (see lsl_st_varan.h)
//[<sd_retval] 0=OK, negative=error (look lsl_st_varan.h)
FUNCTION VIRTUAL GLOBAL VaranManager::ClearDOL
  VAR_INPUT
    ud_dol_type	    	: UDINT;
  END_VAR
  VAR_OUTPUT
    sd_retval		      : DINT;
  END_VAR

  // if there is no VARAN Interface available, we would crash at the call
  if pVaran = NIL then
    sd_retval := VARANMANAGER_DRIVER_NOT_EXISTS;
    return;
  end_if;

  sd_retval := VARAN_iClearDOL( uiManager		:= VaranManagerNr
                              , uiDOLType 	:= ud_dol_type
                              );

  //look if an error occurs
  if ( sd_retval <> VARANMANAGER_OK ) then
    s_ErrorVaranManager.f_ClearDOL := SetVaranDOError ( sd_Error 		  := sd_retval
                                                      , b_manager_off	:= TRUE
                                                      , b_log			    := TRUE
                                                      );
  end_if;

END_FUNCTION //VIRTUAL GLOBAL VaranManager::ClearDOL

//[#ENGLISH]
//=================================================================================================
//Function to read a direct access data object
//=================================================================================================
//[members]	s_DirectAccessDO	:W/R	:structure for direct access
//[>p_us_position_info]pointer to position info( first byte is length )
//[>ud_address]address to read
//[>ud_length]length of data should read
//[>p_ud_data]variable to get pointer to readed data
//[>ud_type] 0=control area, 1=memory area
//[<sd_retval] 0=OK, negative=error (look lsl_st_varan.h)
FUNCTION VIRTUAL GLOBAL VaranManager::RdDO
  VAR_INPUT
    p_us_position_info	: ^USINT;
    ud_address			    :  UDINT;
    ud_length			      :  UDINT;
    p_ud_data			      : ^UDINT;
    ud_type			      	:  UDINT;
  END_VAR
  VAR_OUTPUT
    sd_retval			      :  DINT;
  END_VAR

  //enable semaphore
  To_Multitask.Wait( p_SemaHandle );

  //clear direct access dol list
  sd_retval := ClearDOL( ud_dol_type := VARAN_DOL_DA );

  //look if an error occurs
  if ( sd_retval <> VARANMANAGER_OK ) then
    s_ErrorVaranManager.f_RdDO := SetVaranDOError	( sd_Error 	:= sd_retval
                                                  , b_manager_off	:= TRUE
                                                  , b_log			:= FALSE
                                                  );
    //disable semaphore
    To_Multitask.Signal( p_SemaHandle );
    return;
  end_if;

  //add data object
  sd_retval := AddRdDO( p_us_position_info  := p_us_position_info
                      , ud_dol_type		      := VARAN_DOL_DA
                      , p_ud_handle		      := ( #s_DirectAccessDO.ud_DOHandle )$^UDINT
                      , ud_address		      := ud_address
                      , ud_length			      := ud_length
                      , p_ud_data			      := p_ud_data
                      , ud_type			        := ud_type
                      );

  //look if an error occurs
  if ( sd_retval <> VARANMANAGER_OK ) then
    s_ErrorVaranManager.f_RdDO := SetVaranDOError( sd_Error 		  := sd_retval
                                                 , b_manager_off	:= TRUE
                                                 , b_log			    := FALSE
                                                 );
    //disable semaphore
    To_Multitask.Signal( p_SemaHandle );
    return;
  end_if;

  //set run status of data object on
  s_DirectAccessDO.ud_DOHandle^.ucCtrlStat 	  := VARAN_DO_CONT_RUN;

  //set number of allowed retries
  s_DirectAccessDO.ud_DOHandle^.ucRetrys		  := VM_ALLOWED_RETRIES;

  //set time for retry timeout
  s_DirectAccessDO.ud_DOHandle^.uiRetryTimeout:= VM_RETRY_TIMEOUT_DA + ( ( p_us_position_info^ - 1 ) * VM_HUB_DELAY_TIME );

  //Execute dol
  sd_retval := ExecuteDOL( ud_dol_type := VARAN_DOL_DA );//or VARAN_DOL_EXECUTE_WAIT );

  //look if an error occurs
  if ( sd_retval <> VARANMANAGER_OK ) then
    s_ErrorVaranManager.f_RdDO := SetVaranDOError( sd_Error 		  := sd_retval
                                                 , b_manager_off	:= TRUE
                                                 , b_log			    := FALSE
                                                 );
  end_if;

  //disable semaphore
  To_Multitask.Signal( p_SemaHandle );

END_FUNCTION //VIRTUAL GLOBAL VaranManager::RdDO

//[#ENGLISH]
//=================================================================================================
//Function to write a direct access data object
//=================================================================================================
//[members]	s_DirectAccessDO	:W/R	:structure for direct access
//[>p_us_position_info]pointer to position info( first byte is length)
//[>ud_address]address to write
//[>ud_length]length of data should be written
//[>p_ud_data]pointer to data should be written
//[>ud_type]0=control area, 1=memory area
//[<sd_retval] 0=OK, negative=error (look lsl_st_varan.h)
FUNCTION VIRTUAL GLOBAL VaranManager::WrDO
  VAR_INPUT
    p_us_position_info	: ^USINT;
    ud_address	    		:  UDINT;
    ud_length			      :  UDINT;
    p_ud_data			      : ^UDINT;
    ud_type				      :  UDINT;
  END_VAR
  VAR_OUTPUT
    sd_retval			      :  DINT;
  END_VAR

  //enable semaphore
  To_Multitask.Wait( p_SemaHandle );

  //clear direct access dol list
  sd_retval := ClearDOL( ud_dol_type := VARAN_DOL_DA );

  //look if an error occurs
  if ( sd_retval <> VARANMANAGER_OK ) then
    s_ErrorVaranManager.f_WrDO := SetVaranDOError( sd_Error 		  := sd_retval
                                                 , b_manager_off	:= TRUE
                                                 , b_log			    := FALSE
                                                 );
    //disable semaphore
    To_Multitask.Signal( p_SemaHandle );
    return;
  end_if;

  //add data object
  sd_retval := AddWrDO	( p_us_position_info  := p_us_position_info
                        , ud_dol_type		      := VARAN_DOL_DA
                        , p_ud_handle		      := ( #s_DirectAccessDO.ud_DOHandle )$^UDINT
                        , ud_address		      := ud_address
                        , ud_length			      := ud_length
                        , p_ud_data			      := ( #s_DirectAccessDO.p_ud_DOWrite )$^UDINT
                        , ud_type			        := ud_type
                        );

  //look if an error occurs
  if ( sd_retval <> VARANMANAGER_OK ) then
    s_ErrorVaranManager.f_WrDO := SetVaranDOError( sd_Error 		  := sd_retval
                                                 , b_manager_off	:= TRUE
                                                 , b_log			    := FALSE
                                                 );
    //disable semaphore
    To_Multitask.Signal( p_SemaHandle );
    return;
  end_if;

  //set run status of data object on
  s_DirectAccessDO.ud_DOHandle^.ucCtrlStat 	  := VARAN_DO_CONT_RUN;

  //set number of allowed retries
  s_DirectAccessDO.ud_DOHandle^.ucRetrys		  := VM_ALLOWED_RETRIES;

  //set time for retry timeout
  s_DirectAccessDO.ud_DOHandle^.uiRetryTimeout:= VM_RETRY_TIMEOUT_DA + ( ( p_us_position_info^ - 1 ) * VM_HUB_DELAY_TIME );

  //copy write data to dpram space of data object
  To_StdLib.MemCpy( dest 		:= s_DirectAccessDO.p_ud_DOWrite
                  , source 	:= p_ud_data
                  , size 		:= ud_length
                  );

  //Execute dol
  sd_retval := ExecuteDOL( ud_dol_type := VARAN_DOL_DA );//or VARAN_DOL_EXECUTE_WAIT );

  //look if an error occurs
  if ( sd_retval <> VARANMANAGER_OK ) then
    s_ErrorVaranManager.f_WrDO := SetVaranDOError( sd_Error 		  := sd_retval
                                                 , b_manager_off	:= TRUE
                                                 , b_log			    := FALSE
                                                 );
  end_if;

  //disable semaphore
  To_Multitask.Signal( p_SemaHandle );

END_FUNCTION //VIRTUAL GLOBAL VaranManager::WrDO

//[#ENGLISH]
//=================================================================================================
//Function to get Pll - Time of VaranManager
//=================================================================================================
//[members]	s_VMFunctions		:R/W	:structure for HwControl class
//[<ud_varan_time]varan time in ns
FUNCTION VIRTUAL GLOBAL VaranManager::GetVaranTime
  VAR_INPUT
    p_ud_IsoStartPoint	: ^UDINT;
  END_VAR
  VAR_OUTPUT
    ud_varan_time		    :  UDINT;
  END_VAR

  //if we have no Pll-Time yet
  if ( s_VMFunctions.ud_VaranTime = 0 ) then

    //we must init VaranManager first
    if ( s_VaranManagerSettings.us_InitCounter = 0 ) then
      bExternalInit := true;
      Init();
    end_if;
  end_if;

  ud_varan_time := s_VMFunctions.ud_VaranTime;

  //get iso startpoint to calculate the correct offset
  if ( p_ud_IsoStartPoint <> NIL ) then
    p_ud_IsoStartPoint^ := GetIsoStartPoint();
  end_if;

END_FUNCTION //VIRTUAL GLOBAL VaranManager::GetPllTime

//[#ENGLISH]
//=================================================================================================
//Function to send Sync and trigger Watchdog of Varan Bus
//=================================================================================================
//[<sd_retval] 0=OK, negative=error (look lsl_st_varan.h)
FUNCTION VaranManager::TriggerWatchdog
  VAR_OUTPUT
    sd_retval		    : DINT;
  END_VAR

  if b_PayloadSupport &
     pMultiVaran^.udVersion >= VM_MULTIVARAN_VERSION_FULL_PAYLOAD_AVAILABLE  then

    sd_retval := MULTI_VARAN_iTriggerWatchdog(hManagerNodeHandle  := vmNodeHandle
                                            , udWatchdogType      := LSL_WD_TYPE_MANAGER
                                            );
  elsif pVaran then
    sd_retval := VARAN_iTriggerWd( uiManager := VaranManagerNr );
  end_if;

  //if an error occures
  if ( sd_retval <> VARANMANAGER_OK ) then
    s_ErrorVaranManager.f_TriggerWd := SetVaranDOError	( sd_Error 		  := sd_retval
                                                        , b_manager_off	:= TRUE
                                                        , b_log			    := TRUE
                                                        );
    bd_RtLog.WatchdogTriggerFailed := TRUE;
  end_if;

END_FUNCTION //VIRTUAL GLOBAL VaranManager::TriggerWatchdog

//[#ENGLISH]
//=================================================================================================
//Function to extend Handle List
//=================================================================================================
//[servers]	ManagerOn				:W		:marks VaranManager as valid / ok
//[members]	s_RtHandles				:W		:structure to save Handles and thisp for realtime update methodes
//			s_CyHandles				:W		:structure to save Handles and thisp for cyclic update methodes
//			e_ErrorVaranManager		:W		:enum for Error State
//[>ud_dol_type] type of DOL list( Realtime = 3, cyclic = 4 )
FUNCTION VaranManager::ExtendHandleList
  VAR_INPUT
    ud_dol_type 	: UDINT;
    callOptions 	: USINT;
  END_VAR

  //look if an Error occures
  if ( State = _ClassOk ) then

    //--------------------------------------------------------------------------------------------------------------------
    //look which list type we have
    if ( ud_dol_type = VARAN_DOL_ISO ) then
      IF callOptions AND CALL_OPTION_RT_PRESCAN THEN
        //set right max handle
        s_RtHandles.ud_MaxHandles += VM_EXTEND_HANDLES;

        //realloc memory for list
        s_RtHandles.p_HandleList$^void := To_StdLib.ReAlloc	( mptr 		:= s_RtHandles.p_HandleList
                                                            , newsize := s_RtHandles.ud_MaxHandles * sizeof( t_s_OneHandle )
                                                            );

        //look if we got memory for our Handle list
        if ( s_RtHandles.p_HandleList ) then

          //set new memory to 0
          To_StdLib.MemSet( dest 	:= s_RtHandles.p_HandleList + ( s_RtHandles.ud_MaxHandles - VM_EXTEND_HANDLES ) * sizeof( t_s_OneHandle )
                          , value := 0
                          , size 	:= VM_EXTEND_HANDLES * sizeof( t_s_OneHandle )
                          );

        else
          //if not give out a TRACE and set Manager off
          State 		  := _MemoryFault;
          ManagerOn 	:= 0;

          // we switch off isochronous task
          TurnOffIsoTask();

          //Log entry
#ifdef HWC_LogValue1
          HWC_LogValue1(this, "@0690 (VaranManager::ExtendHandleList) No Memory for Varan Manager available! (Extend Rt - Handles: {0})", s_RtHandles.ud_MaxHandles);
#endif
        end_if;
      END_IF;

      IF callOptions AND CALL_OPTION_RT_POSTSCAN THEN
        //set right max handle
        s_RtPostScanHandles.ud_MaxHandles += VM_EXTEND_HANDLES;

        //realloc memory for list
        s_RtPostScanHandles.p_HandleList$^void := To_StdLib.ReAlloc	( mptr 		:= s_RtPostScanHandles.p_HandleList
                                                                    , newsize := s_RtPostScanHandles.ud_MaxHandles * sizeof( t_s_OneHandle )
                                                                    );

        //look if we got memory for our Handle list
        if ( s_RtPostScanHandles.p_HandleList ) then

          //set new memory to 0
          To_StdLib.MemSet( dest 	:= s_RtPostScanHandles.p_HandleList + ( s_RtPostScanHandles.ud_MaxHandles - VM_EXTEND_HANDLES ) * sizeof( t_s_OneHandle )
                          , value := 0
                          , size 	:= VM_EXTEND_HANDLES * sizeof( t_s_OneHandle )
                          );

        else
          //if not give out a TRACE and set Manager off
          State 		  := _MemoryFault;
          ManagerOn 	:= 0;

          // we switch off isochronous task
          TurnOffIsoTask();

          //Log entry
#ifdef HWC_LogValue1
          HWC_LogValue1(this, "@0023 (VaranManager::ExtendHandleList) No Memory for Varan Manager available! (Extend RtPostScan - Handles: {0})", s_RtPostScanHandles.ud_MaxHandles);
#endif
        end_if;
      END_IF;

    //--------------------------------------------------------------------------------------------------------------------
    elsif ( ud_dol_type = VARAN_DOL_ASY ) then

      //set right max handle
      s_CyHandles.ud_MaxHandles += VM_EXTEND_HANDLES;

      //realloc memory for list
      s_CyHandles.p_HandleList$^void := To_StdLib.ReAlloc	( mptr 		:= s_CyHandles.p_HandleList
                                                          , newsize := s_CyHandles.ud_MaxHandles * sizeof( t_s_OneHandle )
                                                          );

      //look if we got memory for our Handle list
      if ( s_CyHandles.p_HandleList ) then

        //set new memory to 0
        To_StdLib.MemSet( dest 	:= s_CyHandles.p_HandleList + ( s_CyHandles.ud_MaxHandles - VM_EXTEND_HANDLES ) * sizeof( t_s_OneHandle )
                        , value := 0
                        , size 	:= VM_EXTEND_HANDLES * sizeof( t_s_OneHandle )
                        );

      else
        //if not give out a TRACE and set Manager off
        State 		  := _MemoryFault;
        ManagerOn 	:= 0;

        // we switch off isochronous task
        TurnOffIsoTask();

        //Log entry
#ifdef HWC_LogValue1
        HWC_LogValue1(this, "@069A (VaranManager::ExtendHandleList) No Memory for Varan Manager available! (Extend Cy - Handles: {0})", s_CyHandles.ud_MaxHandles);
#endif
      end_if;
    end_if;
  end_if;

END_FUNCTION // VaranManager::ExtendHandleList

//[#ENGLISH]
//=================================================================================================
//Function to call Realtime update methode of a varan class
//=================================================================================================
//[>p_this]Thispointer of Varan_Base class
FUNCTION  VaranManager::CallUpdateRt
  VAR_INPUT
    p_this		  	: p_VaranBase;
  END_VAR

  p_this^.UpdateRt();

END_FUNCTION // VaranManager::CallUpdateRt

//[#ENGLISH]
//=================================================================================================
//Function to call Cyclic update methode of a varan class
//=================================================================================================
//[>p_this]Thispointer of Varan_Base class
FUNCTION  VaranManager::CallUpdateCy
  VAR_INPUT
    p_this		  	: p_VaranBase;
  END_VAR

  p_this^.UpdateCy();

END_FUNCTION // VaranManager::CallUpdateCy

//[#ENGLISH]
//=================================================================================================
//Function to set Error in VaranManager
//=================================================================================================
//[members]	e_ErrorVaranManager		:W		:Enum for Error State
//[>sd_Error]Error of VaranManager
//[>b_manager_off]0=run, 1=set VaranManagerOff
//[>b_log]0=no logging, 1=log fault
FUNCTION  VaranManager::SetVaranDOError
  VAR_INPUT
    sd_error		    : DINT;
    b_manager_off	  : BOOL;
    b_log			      : BOOL;
  END_VAR
  VAR_OUTPUT
    sd_enum_error	  : t_e_VaranErrors;
  END_VAR

  case ( sd_Error ) of

    VARANMANAGER_DRIVER_NOT_EXISTS:         sd_enum_error := _VaranDriverNotExists;
    VARANMANAGER_DOL_TYPE_WRONG:            sd_enum_error := _WrongDOLType;
    VARANMANAGER_RUN_STATUS_WRONG:          sd_enum_error := _WrongRunStatus;
    VARANMANAGER_DO_HANDLE_INVALID:         sd_enum_error := _DOHandleInvalid;
    VARANMANAGER_DO_RAM_FULL:               sd_enum_error := _DORamFull;
    VARANMANAGER_DO_CMD_INVALID:            sd_enum_error := _DOCmdInvalid;
    VARANMANAGER_MANAGER_NOT_EXISTS:        sd_enum_error := _ManagerNotExists;
    VARANMANAGER_DOL_ADDRESS_INVALID:       sd_enum_error := _DOLAddressInvalid;
    VARANMANAGER_UNKNOWN_COMMAND:           sd_enum_error := _UnknownCommand;
    VARANMANAGER_COMPONENT_NOT_EXISTS:      sd_enum_error := _ComponentNotExists;
    VARANMANAGER_CLIENT_NOT_EXISTS:         sd_enum_error := _ClientNotExists;
    VARANMANAGER_CDIAS_EEPROM_NOT_EXISTS:   sd_enum_error := _CdiasEEPromNotExists;
    VARANMANAGER_CDIAS_EEPROM_NO_GRANT:     sd_enum_error := _CdiasEEPromNoGrant;
    VARANMANAGER_CDIAS_EEPROM_NACK:         sd_enum_error := _CdiasEEPromNack;
    VARANMANAGER_PORT_NOT_EXISTS:           sd_enum_error := _PortNotExists;
    VARANMANAGER_PORT_IS_UPLINK:            sd_enum_error := _PortIsUplink;
    VARANMANAGER_PORT_NO_LINK:              sd_enum_error := _PortNoLink;
    VARANMANAGER_NO_MUTEX:                  sd_enum_error := _NoMutex;
    VARANMANAGER_NO_TASK:                   sd_enum_error := _NoTask;
    VARANMANAGER_ID_NOT_FOUND:              sd_enum_error := _IDNotFound;
    VARANMANAGER_ID_NOT_INITIALIZED:        sd_enum_error := _IDNotInitialized;
    VARANMANAGER_INVALID_DEVICE_ADDRESS:    sd_enum_error := _InvalidDeviceAddress;
    VARANMANAGER_CALLBACK_NOT_HANDLED:      sd_enum_error := _CallbackNotHandled;
    VARANMANAGER_NO_MEM:                    sd_enum_error := _NoMem;
    VARANMANAGER_NO_LEGACY_WD:              sd_enum_error := _NoLegacyWd;
    VARANMANAGER_ADMIN_DOL_EXECUTION_ERROR: sd_enum_error := _AdminDOLExecutionError;
    VARANMANAGER_DA_DOL_EXECUTION_ERROR:    sd_enum_error := _DADOLExecutionError;
    VARANMANAGER_SPI_FLASH_NO_ACCESS:       sd_enum_error := _SPIFlashNoAccess;
    VARANMANAGER_CLIENT_NOT_READY:          sd_enum_error := _ClientNotready;
    VARANMANAGER_CLIENT_DISABLED:           sd_enum_error := _ClientDisabled;
    VARANMANAGER_CLIENT_CANT_ENABLE:        sd_enum_error := _ClientCantEnable;
    VARANMANAGER_CDIAS_ADDRESS_INVALID:     sd_enum_error := _CdiasAddressInvalid;
    VARANMANAGER_SPI_FLASH_INVALID:         sd_enum_error := _SPIFlashInvalid;
    VARANMANAGER_SPI_DOL_ID_INVALID:        sd_enum_error := _SPIDOLIDInvalid;
    VARANMANAGER_SPI_DOL_INVALID:           sd_enum_error := _SPIDOLInvalid;
    VARANMANAGER_SPI_REQUIRED_LIST_ERROR:   sd_enum_error := _SPIRequiredListError;
    VARANMANAGER_SPI_CHKSUM_ERROR:          sd_enum_error := _SPIChksumError;
    VARANMANAGER_PARAMETER_INVALID:         sd_enum_error := _ParameterInvalid;
    VARANMANAGER_DO_TYPE_NOT_SUPPORTED:     sd_enum_error := _DOTypeNotSupported;
    VARANMANAGER_DMA_ERROR:                 sd_enum_error := _DMAError;
    VARANMANAGER_PROPERTY_ID_INVALID:       sd_enum_error := _PropertyIDInvalid;
    VARANMANAGER_PROPERTY_VALUE_INVALID:    sd_enum_error := _PropertyValueInvalid;
    VARANMANAGER_DO_NUMBER_OVERFLOW:        sd_enum_error := _DONumberOverflow;
    VARANMANAGER_API_USAGE_NOT_ALLOWED:     sd_enum_error := _APIUsageNotAllowed;
    VARANMANAGER_NODE_TYPE_WRONG:           sd_enum_error := _NodeTypeWrong;
    VARANMANAGER_DATA_LENGTH_INVALID:       sd_enum_error := _DataLengthInvalid;
    VARANMANAGER_DO_TYPE_INVALID:           sd_enum_error := _DOTypeInvalid;
    VARANMANAGER_OPERATION_NOT_ALLOWED:     sd_enum_error := _OperationNotAllowed;
    VARANMANAGER_NODE_NUMBER_OVERFLOW:      sd_enum_error := _NodeNumberOverflow;
    VARANMANAGER_NO_HANDLE_FOUND:           sd_enum_error := _NoHandleFound;

    -2147482560:                            sd_enum_error := _TimeoutVaran;  //16#8000_0440

  else
    if sd_Error < 0 then
      sd_enum_error := _UnknownFault;
    end_if;
  end_case;

  s_VaranManagerSettings.sd_LastError 	:= sd_error;
  s_ErrorVaranManager.ud_ErrorCounter   += 1;

  //Log entry
  if b_log then
#ifdef HWC_LogValue1
    HWC_LogValue1(this, "@06A4 (VaranManager::SetVaranDOError) Error happened with ErrorCode {0}", s_VaranManagerSettings.sd_LastError$UDINT);
#endif
  end_if;

  //should we set VaranManager off
  if ( b_manager_off = TRUE ) then

    //Log entry
    if b_log then
#ifdef HWC_LogError
      HWC_LogError(this, "@06AE (VaranManager::SetVaranDOError) Is set off because of last Error!");
#endif
    end_if;

    ManagerOn 		:= 0;

    // End the PostInit Phase as it can't be ended regularly as the VM is set off.
    // Otherwise PostInit Phase would end on timeout.
    bPostInitModulesReady := TRUE;

    //to make log entry in cyclic
    s_VaranManagerSettings.b_LogError := TRUE;

    // we switch off isochronous task
    TurnOffIsoTask();

    //set Hw off
    To_HwControl.SetHardwareOff( e_error := State );

    State 			:= sd_enum_error;
  end_if;

END_FUNCTION // VaranManager::SetVaranDOError

//[#ENGLISH]
//=================================================================================================
//Function to get µs time
//=================================================================================================
//[<ud_us_sec(EAX)]µs - Time
FUNCTION  VaranManager::GetMuSec
  VAR_OUTPUT
    ud_us_sec(EAX)		: UDINT;
  END_VAR

#ifdef _LSL_TARGETARCH_X86
  SAVE_REG();
#endif
  ud_us_sec := OS_ReadMicroSec();
#ifdef _LSL_TARGETARCH_X86
  RESTORE_REG();
#endif

END_FUNCTION // VaranManager::GetMuSec

//[#ENGLISH]
//=================================================================================================
//Function to get Varan class position in a string
//=================================================================================================
//[>p_us_info] pointer to save position info (first byte is length)
//[<sd_retval]0=OK, -1=to many hubs( max.15 )
#pragma warning(disable: 73)
FUNCTION VIRTUAL GLOBAL VaranManager::GetVaranPosition
  VAR_INPUT
    p_us_info	  	: ^USINT;
  END_VAR
  VAR_OUTPUT
    sd_retval	  	:  DINT;
  END_VAR

  //I am the Manager -> do nothing
  sd_retval := -1;

END_FUNCTION //VIRTUAL GLOBAL VaranManager::GetVaranPosition
#pragma warning(default: 73)
//[#ENGLISH]
//=================================================================================================
//Function to install callback function for hot plug and play
//=================================================================================================
//[>p_us_position_info]pointer to position info( first byte is length)
//[>ud_action_ptr]pointer to function
//[>ud_thisp]thispointer
//[>sd_required]is class required
FUNCTION VIRTUAL GLOBAL VaranManager::SetObjectCallback
  VAR_INPUT
    p_us_position_info	: ^USINT;
    ud_action_ptr	    	:  UDINT;
    ud_thisp			      :  UDINT;
    sd_required		    	:  DINT;
  END_VAR
  VAR_OUTPUT
    sd_retval		        :  DINT;
  END_VAR
  VAR
    p_one_module        : ^p_VaranBase;
    p_one_posstring     : ^pVoid;
  END_VAR

  sd_retval := AddObjectCallback( p_us_position_info:=p_us_position_info
                                , ud_action_ptr:= ud_action_ptr
                                , ud_thisp:= ud_thisp
                                , sd_required:= sd_required
                                );

  // don't save the this pointer of the varan manager itself
  if p_us_position_info then
    // save pthis to internal list
    if ( s_ModuleList.ud_NrOfModules = s_ModuleList.ud_MaxModules ) then

      //extend list
      sd_retval := ExtendModuleList();

      //if an error occured return
      if ( sd_retval <> VARANMANAGER_OK ) then
        s_ErrorVaranManager.f_SetObjectCallback := SetVaranDOError	( sd_Error 		  := sd_retval
                                                                    , b_manager_off	:= TRUE
                                                                    , b_log			    := TRUE
                                                                    );
        return;
      end_if;
    end_if;

    //set pointer to next free handle entry
    p_one_module 	    := (s_ModuleList.p_ModuleList + ( s_ModuleList.ud_NrOfModules * sizeof( p_VaranBase ) ))$^p_VaranBase;
    p_one_module^	    := ud_thisp$p_VaranBase;

    //set pointer to next free handle entry
    p_one_posstring 	:= (s_ModuleList.p_PositionList + ( s_ModuleList.ud_NrOfModules * sizeof(pVoid) ))$^pVoid;
    p_one_posstring^	:= p_us_position_info$^pVoid;

    //increase number of handles
    s_ModuleList.ud_NrOfModules += 1;
  end_if;

END_FUNCTION //VIRTUAL GLOBAL VaranManager::SetObjectCallback

//[#ENGLISH]
//=================================================================================================
//Function sets Manager off
//=================================================================================================
//[server]	ManagerOn			:W		:state of Manager (On/Off)
//[members]	s_DirectAccessDO		:W/R	:structure for direct access
//			s_VaranManagerSettings	:W		:structure for different varan settings
//[>e_error]reason why varan Manager is set off
FUNCTION VIRTUAL GLOBAL VaranManager::SetManagerOff
  VAR_INPUT
    e_error		: t_e_VaranErrors;
  END_VAR
  VAR
    i         : UDINT;
    pHelp     : ^p_VaranBase;
  END_VAR

  ManagerOn 	:= 0;

  // we switch off isochronous task
  TurnOffIsoTask();

  if ( State = _ClassOk ) then
    State		:= e_error;

    //to make log entry in cyclic
    s_VaranManagerSettings.b_LogError := TRUE;

    //update state of modules connected befor error
    if ( s_ModuleList.ud_NrOfModules > 0 ) then

      //check all connected classes
      pHelp := s_ModuleList.p_ModuleList;
      for i := 0 to s_ModuleList.ud_NrOfModules - 1 do

        if pHelp^^.State = _ClassOk then
          //module was connected before Manager was turned off, set new state
          pHelp^^.State   := _ModuleFoundButManagerIsOff;
          pHelp^^.Online  := 0; // also reset the online server
        end_if;

        //get pointer on next handle
        pHelp += sizeof(p_VaranBase);
      end_for;
    end_if;
  end_if;

  //set HwControl off
  To_HwControl.SetHardwareOff( e_error := e_error );

  // End the PostInit Phase as it can't be ended regularly as the VM is set off.
  // Otherwise PostInit Phase would end on timeout.
  bPostInitModulesReady := TRUE;

END_FUNCTION //VIRTUAL GLOBAL VaranManager::SetManagerOff

//[#ENGLISH]
//=================================================================================================
//Function set a varan error
//=================================================================================================
//[members]	s_VaranManagerSettings	:W		:structure for different varan settings
//[locals]	p_handle	:W/R	:pointer to a varan handle
//			p_data		:W/R	:pointer to data of data object
//			sd_retval	:W/R	:return value of OS - functions
//[>p_Node]pointer to Node string
FUNCTION VIRTUAL GLOBAL VaranManager::SetVaranError
  VAR_INPUT
    p_Node		: ^USINT;
  END_VAR
  VAR
    p_handle	: ^LSL_VARANFRAME;
    p_data		: ^UDINT;
    sd_retval	:  DINT;
    NodeHandle:  UDINT;
  END_VAR

  p_Handle 	:= NIL;
  p_Data 		:= NIL;

  //look if init was executed
  if ( s_VaranManagerSettings.us_InitCounter = 0 ) then
    bExternalInit := true;
    Init();
  end_if;

  //log error if we have one
  if ( s_VaranManagerSettings.b_LogError ) then
    LogError();
  end_if;

  if b_PayloadSupport then

    // see if we can get the handle of the target device
    sd_retval := MULTI_VARAN_iGetNodeHandle(  udManagerNumber := VaranManagerNr
                                           ,  pszHardwarePath := p_Node
                                           ,  phNodeHandle    := #NodeHandle
                                           );

    if sd_retval = VARANMANAGER_OK then
      // we got the current node handle => use it
      MULTI_VARAN_iReportVaranError( diErrorNumber := VM_ERROR_REQUIRED
                                   , hErrorNode    := NodeHandle
                                   );
    else
      // we don't have the current handle => use the manager handle
      MULTI_VARAN_iReportVaranError( diErrorNumber := VM_ERROR_REQUIRED
                                   , hErrorNode    := vmNodeHandle
                                   );
    end_if;

  elsif pVaran then

    //clear DOL list
    sd_retval := VARAN_iClearDOL( uiManager		:= VaranManagerNr
                                , uiDOLType 	:= VARAN_DOL_DA
                                );

    //look for an Error
    if ( sd_retval <> VARANMANAGER_OK ) then
      s_ErrorVaranManager.f_SetVaranError := SetVaranDOError	( sd_Error 		  := sd_retval
                                                              , b_manager_off	:= TRUE
                                                              , b_log			    := FALSE
                                                              );
      return;
    end_if;

    //Install Varan data object
    sd_retval := VARAN_iAddDOToDOL	( uiManager			  := VaranManagerNr
                                    , pucNode			    := p_Node
                                    , uiDOLType 		  := VARAN_DOL_DA
                                    , puiDOHandle		  := ( #p_Handle )$^UDINT
                                    , uiCmd				    := VARAN_CMD_MEMORY_READ
                                    , uiAddressRead		:= 16#1
                                    , uiLengthRead		:= 1
                                    , pucRead			    := ( #p_Data )$^UDINT
                                    , uiAddressWrite	:= 0
                                    , uiLengthWrite		:= 0
                                    , pucWrite			  := NIL
                                    );

    //look for an Error
    if ( sd_retval <> VARANMANAGER_OK ) then
      s_ErrorVaranManager.f_SetVaranError := SetVaranDOError	( sd_Error 		  := sd_retval
                                                              , b_manager_off	:= TRUE
                                                              , b_log			    := FALSE
                                                              );
      return;
    end_if;

    //set run status of data object on
    p_Handle^.ucCtrlStat 	    := VARAN_DO_SINGLE_RUN or VARAN_DO_REQUIRED;
    p_Handle^.uiRetryTimeout  := 1000;
    p_Handle^.ucRetrys 		    := 1;
    p_Handle^.ucRetryCounter  := 0;

    //Execute DOL list
    sd_retval := VARAN_iExecuteDOLDA( uiManager := VaranManagerNr );

    //look for an Error
    if ( sd_retval <> VARANMANAGER_OK ) then
      s_ErrorVaranManager.f_SetVaranError := SetVaranDOError	( sd_Error 		  := sd_retval
                                                              , b_manager_off	:= TRUE
                                                              , b_log			    := FALSE
                                                              );
      return;
    end_if;

  end_if;

END_FUNCTION //VIRTUAL GLOBAL VaranManager::SetVaranError

//[#ENGLISH]
//=================================================================================================
//Function give back a nono second counter value of VaranManager
//=================================================================================================
//[members]	p_ManagerStructure		:W/R	:pointer for manager structure (from OS)
//			s_VaranManagerSettings	:R		:structure for different varan settings
//[<ud_ns_counter]nano second counter value
FUNCTION VIRTUAL GLOBAL VaranManager::GetNsTime
  VAR_OUTPUT
    ud_ns_counter		: UDINT;
  END_VAR

  //look if init was executed
  if ( s_VaranManagerSettings.us_InitCounter = 0 ) then
    bExternalInit := true;
    Init();
  end_if;

  if b_PayloadSupport  &
     pMultiVaran^.udVersion >= VM_MULTIVARAN_VERSION_FULL_PAYLOAD_AVAILABLE then
    MULTI_VARAN_iGetTimeUpCounter( hManagerNodeHandle := vmNodeHandle
                                 , pudTimeUpCounterNs := #ud_ns_counter
                                 );
  elsif ( p_ManagerStructure <> NIL ) then  //if we have the Manager structure

    ud_ns_counter := p_ManagerStructure^.uiTUpCounter;

  end_if;

END_FUNCTION //VIRTUAL GLOBAL VaranManager::GetNsTime

//[#ENGLISH]
//=================================================================================================
//Function trace a Realtime Overlap fault
//=================================================================================================
//[server]	ManagerOn				:W		:state of Manager (On/Off)
//			State					:R		:State of class
//[members]	s_VaranManagerSettings	:W		:structure for different varan settings
FUNCTION  VaranManager::TRACE_RtOverlap

  if ( State = _ClassOk ) then

    State 		:= _TimesliceError;
    ManagerOn	:= 0;

    // we switch off isochronous task
    TurnOffIsoTask();

    s_VaranManagerSettings.b_LogError := TRUE;

    bd_RtLog.TimeSliceError := TRUE;

    //set Hw off
    To_HwControl.SetHardwareOff( e_error := _TimesliceError );
  end_if;

END_FUNCTION // VaranManager::TRACE_RtOverlap

//[#ENGLISH]
//=================================================================================================
//Function to get watchdog or timeslice error
//=================================================================================================
//[server]	ManagerOn				:W		:state of Manager (On/Off)
//			State					:R		:State of class
//[members]	s_VaranManagerSettings	:W		:structure for different varan settings
//[>ud_reason]reason of callback
FUNCTION  VaranManager::Varan_CallBack
  VAR_INPUT
    ud_reason   	: UDINT;
  END_VAR
  VAR
    pHelp         : ^t_s_FlexHub;
    HandleError   : BOOL;
#ifdef VARANMANAGER_CB_VMC_BUF_DA
    Time1, Time2  : UDINT;
#endif
  END_VAR

  if ( State = _ClassOk )
#ifdef VARANMANAGER_CB_VMC_BUF_DA
   | ( ud_reason = VARANMANAGER_CB_VMC_BUF_DA )
#else
  #pragma message("Need newer lsl_st_varan.h file for direct access buffer of vmc");
#endif
    then

    // if we're not told other ways, raise "exception" (time slice error or whatever)
    HandleError := TRUE;

    case ( ud_reason ) of
// **********************************************************************************************************************************************
      VARANMANAGER_CB_TIME_SLICE_ERROR:

#ifdef VARAN_iSetManagerCallbackOnVmcBufDaInt
        if (_RTOSVersion >= VM_DA_BUFFER_AVAILABLE) & pVaran then
          VARAN_iSetManagerCallbackOnVmcBufDaInt(0);
        end_if;
#endif
        State := _TimesliceErrorIRQ;

// **********************************************************************************************************************************************
      VARANMANAGER_CB_WATCHDOG_ERROR:
#ifdef VARAN_iSetManagerCallbackOnVmcBufDaInt
        if (_RTOSVersion >= VM_DA_BUFFER_AVAILABLE) & pVaran then
          VARAN_iSetManagerCallbackOnVmcBufDaInt(0);
        end_if;
#endif
        State := _WatchdogError;

// **********************************************************************************************************************************************
#ifdef VARANMANAGER_CB_VMC_BUF_DA
      VARANMANAGER_CB_VMC_BUF_DA:

Time1 := OS_READMICROSEC();

        // don't raise exception
        HandleError := FALSE;

        // read data from buffer (first byte is irq quit address) and store it in application memory

        // first copy data
        if DA_IRQ_Length > VM_CLIENT_HEADER_SIZE then
          To_Stdlib.MemCpy(dest   := DA_IRQ_pData + VM_CLIENT_HEADER_SIZE
                         , source := p_ManagerClientSpace + VM_CLIENT_DA_RD_OFFSET + VM_CLIENT_HEADER_SIZE
                         , size   := DA_IRQ_Length - VM_CLIENT_HEADER_SIZE
                         );
        end_if;

        // switch buffer and read last(first) 4 Byte (to quit irq after read-out all data)
        DA_IRQ_pData^$UDINT :=  (p_ManagerClientSpace + VM_CLIENT_DA_RD_OFFSET)^$UDINT;

        // call user irq method
        DA_IRQ_pFunc$IRQMethodDummy(DA_IRQ_pthis);

// do not delete time measurement, could be useful when someone waits for a response in the same cycle
Time2 := OS_READMICROSEC();
DAIRQTime := Time2 - Time1;
#endif
// **********************************************************************************************************************************************
      VARANMANAGER_CB_DISCONNECT,
      VARANMANAGER_CB_CONNECT:

        // don't raise exception
        HandleError := FALSE;

      // refresh flex hub classes

        // call all flexhubs
        if pFlexHubs then

          // TODO: check which component has been dis-/connected and store info in t_s_FlexHub_Parameters, which will be passed to the flexhubs

          pHelp := pFlexHubs;
          while pHelp <> NIL do
            WR(pHelp^.pServer, ud_reason$DINT);
            pHelp := pHelp^.pNext;
          end_while;
        end_if;
    end_case;

    if HandleError then
      // only for errors

      //to make log entry in cyclic
      s_VaranManagerSettings.b_LogError := TRUE;

      // we switch off isochronous task
      TurnOffIsoTask();

      //set Hw off
      To_HwControl.SetHardwareOff( e_error := State );

      //set Manager off
      ManagerOn := 0;
    end_if;
  end_if;

END_FUNCTION // VaranManager::Varan_CallBack

//[#ENGLISH]
//=================================================================================================
//Function to get pointer to node information
//=================================================================================================
//[>p_us_position_info]pointer to position info( first byte is length)
//[>p_node_info]pointer to node info
FUNCTION VIRTUAL GLOBAL VaranManager::GetNodeInfo
  VAR_INPUT
    p_us_position_info	: ^USINT;
    p_node_info		    	: ^PLSL_VARANNODEINFO;
  END_VAR
  VAR_OUTPUT
    sd_retval			      :  DINT;
  END_VAR
  VAR
    ud_NodeHandle       : UDINT;
    nodeProperty        : LSL_PROPERTY_VALUE_PAIR;
  END_VAR

  //look if init was executed
  if ( s_VaranManagerSettings.us_InitCounter = 0 ) then
    bExternalInit := true;
    Init();
  end_if;

  if p_us_position_info & p_node_info then
    if b_PayloadSupport then //----------------------------------------------------------------------------------------------------------

      // Check the pointer, the data is now stored to the pointer
      if p_node_info then
        sd_retval := MULTI_VARAN_iGetNodeHandle ( udManagerNumber := VaranManagerNr
                                                , pszHardwarePath := p_us_position_info
                                                , phNodeHandle    := #ud_NodeHandle
                                                );

        // Return the ErrorCode
        if sd_retval <> VARANMANAGER_OK then
          return;
        end_if;

        sd_retval := MULTI_VARAN_iGetNodeInformation( hNodeHandle := ud_NodeHandle
                                                    , psNodeInfo  := p_node_info^
                                                    );
